Staubli VAL3: click_Hold.pgx

program click_Hold()
  local bool l_bResult
begin
   //暂停机器人
  l_bResult=userPageConfirm("确认暂停机器人？")
  if l_bResult
    rs:bToPause=true
    delay(0.2)
    rs:bToPause=false
  endIf
end
